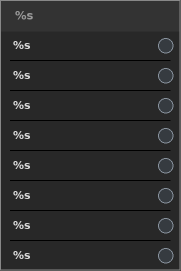
VISUALIZATION FRM_8BitDisplay  // 181x271
VAR_INPUT
   sName: STRING;  

    sBit0: STRING;
    sBit1: STRING;
    sBit2: STRING;
    sBit3: STRING;
    sBit4: STRING;
    sBit5: STRING;
    sBit6: STRING;
    sBit7: STRING; 
   
    bBit0: BOOL;
    bBit1: BOOL;
    bBit2: BOOL;
    bBit3: BOOL;
    bBit4: BOOL;
    bBit5: BOOL;
    bBit6: BOOL;
    bBit7: BOOL;
END_VAR
    Rectangle (0,30 181x241)
    Textfield (10,40 141x11), "%s", text variable: sBit0
    Textfield (10,70 141x11), "%s", text variable: sBit1
    Textfield (10,100 141x11), "%s", text variable: sBit2
    Textfield (10,130 141x11), "%s", text variable: sBit3
    Textfield (10,160 141x11), "%s", text variable: sBit4
    Textfield (10,190 151x11), "%s", text variable: sBit5
    Textfield (10,220 141x11), "%s", text variable: sBit6
    Textfield (10,250 141x11), "%s", text variable: sBit7
    Line (10,60) (170,60)
    Line (10,90) (170,90)
    Line (10,120) (170,120)
    Line (10,150) (170,150)
    Line (10,180) (170,180)
    Line (10,210) (170,210)
    Line (10,240) (170,240)
    Textfield (0,0 181x31), "%s", text variable: sName
    Ellipse (158,38 15x15), colour toggle: bBit0
    Ellipse (158,68 15x15), colour toggle: bBit1
    Ellipse (158,98 15x15), colour toggle: bBit2
    Ellipse (158,128 15x15), colour toggle: bBit3
    Ellipse (158,158 15x15), colour toggle: bBit4
    Ellipse (158,188 15x15), colour toggle: bBit5
    Ellipse (158,218 15x15), colour toggle: bBit6
    Ellipse (158,248 15x15), colour toggle: bBit7
END_VISUALIZATION

(* stored: Version 1.1.0.1
   Visu FRM_8BitDisplay: Id {1eedfe70-0c03-01dd-3302-d09f96606fdf} *)
